GLOBALCONSTANTS DiagCodes (* PLCopen Safety Part 1 Ch. 5.2 - generic DiagCode shared by all SF_ blocks *)
  (* Standard: 61499-1; Description: Copyright (c) 2026 Meisterschulen am Ostbahnhof This program and the accompanying materials are made available under the terms of the Eclipse Public License 2.0 which is available at https://www.eclipse.org/legal/epl-2.0/ SPDX-License-Identifier: EPL-2.0 *)
  (* Version 2.0, 2026-10-09, Franz Höpfinger, Meisterschulen am Ostbahnhof, Split into DiagCodes (generic, Ch. 5.2) + ResetButtonDiagCodes + EmergencyStopDiagCodes (FB-specific, Ch. 6.x.6). Previously held every code in one file. *)
  (* Version 1.0, 2026-10-09, Franz Höpfinger, Meisterschulen am Ostbahnhof, Source: PLCopen TC5 Safety Part 1, Version 2.10, Chapter 6.1.6 DiagCode table. *)
  PACKAGE logiBUS::safety::PLCopen::const;
  VAR_GLOBAL CONSTANT
    IDLE : WORD := 16#0000; (* 0000 - FB not active, generic for all SF_ blocks *)
  END_VAR
END_GLOBALCONSTANTS
